FUNCTION_BLOCK AutomaticExtractionHandler_Test EXTENDS TcUnit.FB_TestSuite
VAR_INPUT
END_VAR
VAR_OUTPUT
END_VAR
VAR
END_VAR


// Control valve calibration tests

// Manual mode tests
(*
-State must be MANUAL_EXTRACTION when automatic extraction not commanded
-State must be MANUAL_EXTRACTION when calibration is not done (even if automatic extraction started)
-All valves must be closed when manual extraction entered
-Inlet and outlet valve signals must reflect the command during manual extraction
-Internal calibration start command must be false during manual extraction
-Pumping pressure decrease command must be false during manual extraction
*)
manualModeTests();
// Automatic mode tests
(*
-State must not be MANUAL_EXTRACTION when automatic extraction commanded
-extractiveOutOnOffValveCommand should be opposite to stateMachines co2onOffValveClosed output
-controlValveOpeningPercentage should be the same as commanded by StateMachine
-If reactor filling not active, reactor outlet valve should remain closed
-If reactor filling active, pressure reference should be updated
-If reactor filling active, reactor outlet valve should be open if outlet valve commands it to
*)
automaticModeTests();

METHOD automaticModeTests
VAR
	handler : AutomaticExtractionHandler;
	testParams : ST_AutomaticExtractionHandlerTest;
END_VAR

TEST('1: State must not be MANUAL_EXTRACTION when automatic extraction commanded and calibration done');

    handler(
		startAutomaticExtraction := TRUE,
		calibrateDone := TRUE);

    AssertEquals_BOOL(
        Expected := FALSE,
        Actual := (handler.automaticExtractionState = E_AutomaticExtractionState.MANUAL_EXTRACTION
        ),
        Message := 'State MANUAL_EXTRACTION when automatic extraction commanded and calibration done'
    );

TEST_FINISHED();

TEST('2: extractiveOutOnOffValveCommand should be opposite to stateMachines co2onOffValveClosed output');

	handler.setTestMode(
		testParams := testParams,
		reset := TRUE);    

	handler(
		startAutomaticExtraction := TRUE,
		calibrateDone := TRUE);

    AssertEquals_BOOL(
        Expected := TRUE,
        Actual := (handler.extractiveOutOnOffValveAutoCommand
        ),
        Message := 'extractiveOutOnOffValveCommand should be opposite to stateMachines co2onOffValveClosed output'
    );

TEST_FINISHED();
END_METHOD

METHOD manualModeTests : BOOL
VAR
	handler : AutomaticExtractionHandler;
	testParams : ST_AutomaticExtractionHandlerTest;
END_VAR

TEST('1: State must be MANUAL_EXTRACTION when automatic extraction not commanded');

    handler();

    AssertEquals_BOOL(
        Expected := TRUE,
        Actual := (handler.automaticExtractionState = E_AutomaticExtractionState.MANUAL_EXTRACTION
        ),
        Message := 'State not MANUAL_EXTRACTION when automatic extraction not commanded'
    );

TEST_FINISHED();

TEST('2: State must be MANUAL_EXTRACTION when calibration is not done (even if automatic extraction started');

	handler.setTestMode(
					testParams := testParams,
					reset := TRUE);

    handler(
		startAutomaticExtraction := TRUE,
		calibrateDone := FALSE);

    AssertEquals_BOOL(
        Expected := TRUE,
        Actual := (handler.automaticExtractionState = E_AutomaticExtractionState.MANUAL_EXTRACTION
        ),
        Message := 'State not MANUAL_EXTRACTION when calibration unfinished'
    );

TEST_FINISHED();

TEST('3: All valves must be closed when manual extraction entered');

	handler.setTestMode(
					testParams := testParams,
					reset := TRUE);

    handler(
		startAutomaticExtraction := FALSE,
		calibrateDone := FALSE);

    AssertEquals_BOOL(
        Expected := FALSE,
        Actual := (handler.reactorInletValve OR handler.reactorOutletValve ),
        Message := 'All valves not closed when manual extraction entered'
    );

TEST_FINISHED();

TEST('4: Inlet and outlet valve signals must reflect the command during manual extraction');

	handler.setTestMode(
					testParams := testParams,
					reset := TRUE);

    handler(
		startAutomaticExtraction := FALSE,
		slurryInValveCommand := TRUE,
		slurryOutValveCommand := TRUE,
		calibrateDone := FALSE);

    AssertEquals_BOOL(
        Expected := TRUE,
        Actual := (handler.reactorOutletValve AND handler.reactorInletValve),
        Message := 'Inlet and outlet valve signals not reflecting the command during manual extraction'
    );

TEST_FINISHED();

TEST('5: Internal calibration start command must be false during manual extraction');

	handler.setTestMode(
					testParams := testParams,
					reset := TRUE);

    handler();

    AssertEquals_BOOL(
        Expected := FALSE,
        Actual := handler.startCalibration,
        Message := 'Internal calibration start command not false during manual extraction'
    );

TEST_FINISHED();

TEST('6: Pumping pressure decrease command must be false during manual extraction');

	handler.setTestMode(
					testParams := testParams,
					reset := TRUE);

    handler();

    AssertEquals_BOOL(
        Expected := FALSE,
        Actual := handler.decreasePumpSetpoint,
        Message := 'Pumping pressure decrease command not false during manual extraction'
    );

TEST_FINISHED();
END_METHOD

END_FUNCTION_BLOCK

(* stored: Version 1.1.0.1, ProductVersion 3.1.4024.9
   POU AutomaticExtractionHandler_Test: Id {3293b6f1-72e0-4bd1-a306-0636ecf992c0}, SpecialFunc None
   Method automaticModeTests: Id {3efe2a47-b026-479c-ba62-fb8061c61cc0}
   Method manualModeTests: Id {77cb51b6-87c0-4878-89fc-f556f6bc106a} *)
